// TIA Portal V19 export
TYPE "ST_EMG"
   STRUCT
      EMG_1 : Bool;
      EMG_BT : Bool;
      EMG_ControlPanel : Bool;
      EMG_Robot_1 : Bool;
      EMG_Robot_2 : Bool;
      EMG_Robot_3 : Bool;
      EMG_7 : Bool;
      EMG_8 : Bool;
      EMG_9 : Bool;
      EMG_10 : Bool;
      EMG_11 : Bool;
      EMG_12 : Bool;
      EMG_13 : Bool;
      EMG_14 : Bool;
      EMG_General : Bool;
   END_STRUCT;
END_TYPE
